// Hour-angle-axis correction (degrees) for a cross-declination offset on the sky (fHourAngleOffset, degrees) at
// declination fDeclination (degrees): fHourAngleOffset / COS(fDeclination). Near the pole 1/COS grows without bound
// and is a division by zero at +-90 deg, so COS is floored at COS(89.5 deg) (factor 115 at most) and the result is
// limited to +-10 deg, the bound BROTLib puts on the offset command (BROTLib#27, same as MONETcommon's
// F_AzimuthOffsetOnAxis near the zenith). Below |dec| = 89.5 deg the result is unchanged.
FUNCTION F_HourAngleOffsetOnAxis : LREAL
VAR_INPUT
	fHourAngleOffset	: LREAL;	// cross-declination offset on the sky, degrees
	fDeclination		: LREAL;	// declination, degrees
END_VAR
VAR CONSTANT
	D2R				: LREAL := 0.017453292519943295;
	MIN_COS			: LREAL := 0.008726535498373935;	// COS(89.5 deg)
	MAX_AXIS_OFFSET	: LREAL := 10.0;					// degrees
END_VAR

F_HourAngleOffsetOnAxis := LIMIT(-MAX_AXIS_OFFSET, fHourAngleOffset / MAX(COS(fDeclination * D2R), MIN_COS), MAX_AXIS_OFFSET);

END_FUNCTION

(* stored: Version 1.1.0.1, ProductVersion 3.1.4024.15
   POU F_HourAngleOffsetOnAxis: Id {6b5752f8-ec6b-4668-ba5b-468b73dcd36c}, SpecialFunc None *)
